Fanuc KAREL source: KT00473.KL

PROGRAM KT00473
%NOLOCKGROUP
VAR
  P1: POSITION
  P2: POSITION
  OUT: BOOLEAN
BEGIN
  OUT = P1 >=< P2
END KT00473
